// TIA Portal V20 export
// export: Created 2026-10-12T05:42:35.0167656Z, ExportSetting WithDefaults, DisplayName Totally Integrated Automation Portal, DisplayVersion V20, DisplayName TIA Portal Openness, DisplayVersion V20, DisplayName TIA Portal Teamcenter Gateway, DisplayVersion V20, DisplayName TIA Portal Version Control Interface, DisplayVersion V20, DisplayName SINAMICS Startdrive Advanced, DisplayVersion V20 SP1 Update 2, DisplayName SINAMICS Startdrive G110M, G120, G120C, G120D, G120P, G115D, DisplayVersion V20 SP1 Update 2, DisplayName SINAMICS Startdrive G130, G150, S120, S150, SINAMICS MV, G220, S200, S210, DisplayVersion V20 SP1 Update 2, DisplayName STEP 7 Professional, DisplayVersion V20, DisplayName STEP 7 Safety, DisplayVersion V20, DisplayName WinCC Basic/Comfort/Advanced, DisplayVersion V20, DisplayName WinCC Professional, DisplayVersion V20, DisplayName WinCC Unified, DisplayVersion V20
FUNCTION_BLOCK "FB_LD_PressDemoHome"   // FB7, LAD
{ S7_Optimized_Access := 'TRUE' }
VERSION : 0.1
// stored: AutoNumber true, IsIECCheckEnabled false, IsRetainMemResEnabled false, MemoryReserve 100, SetENOAutomatically false, UDAEnableTagReadback false
   VAR_INPUT
      Run { ExternalWritable := 'False'} : Bool;
      Reset { ExternalWritable := 'False'} : Bool;
      OwnerIndex { ExternalWritable := 'False'} : DInt;
      Delta { ExternalWritable := 'False'} : Time;
   END_VAR
   VAR_IN_OUT
      PressRam : "FB_CylinderCM";
      Door : "FB_CylinderCM";
      PartSlide : "FB_CylinderCM";
   END_VAR
   VAR
      Seq { ExternalWritable := 'False'} : "FRK_SequenceCtx";
      Row1 { ExternalWritable := 'False'} : "FRK_SequenceRow";
      Row2 { ExternalWritable := 'False'} : "FRK_SequenceRow";
      Row3 { ExternalWritable := 'False'} : "FRK_SequenceRow";
      Row4 { ExternalWritable := 'False'} : "FRK_SequenceRow";
      At0 { ExternalAccessible := 'False'; ExternalVisible := 'False'; ExternalWritable := 'False'} : Bool;
      At900 { ExternalAccessible := 'False'; ExternalVisible := 'False'; ExternalWritable := 'False'} : Bool;
      At910 { ExternalAccessible := 'False'; ExternalVisible := 'False'; ExternalWritable := 'False'} : Bool;
      At999 { ExternalAccessible := 'False'; ExternalVisible := 'False'; ExternalWritable := 'False'} : Bool;
      Ready1 { ExternalAccessible := 'False'; ExternalVisible := 'False'; ExternalWritable := 'False'} : Bool;
      Ready2 { ExternalAccessible := 'False'; ExternalVisible := 'False'; ExternalWritable := 'False'} : Bool;
      Ready3 { ExternalAccessible := 'False'; ExternalVisible := 'False'; ExternalWritable := 'False'} : Bool;
      Ready4 { ExternalAccessible := 'False'; ExternalVisible := 'False'; ExternalWritable := 'False'} : Bool;
      Ready5 { ExternalAccessible := 'False'; ExternalVisible := 'False'; ExternalWritable := 'False'} : Bool;
      Advance { ExternalAccessible := 'False'; ExternalVisible := 'False'; ExternalWritable := 'False'} : Bool;
   END_VAR
BEGIN

REGION Network 1
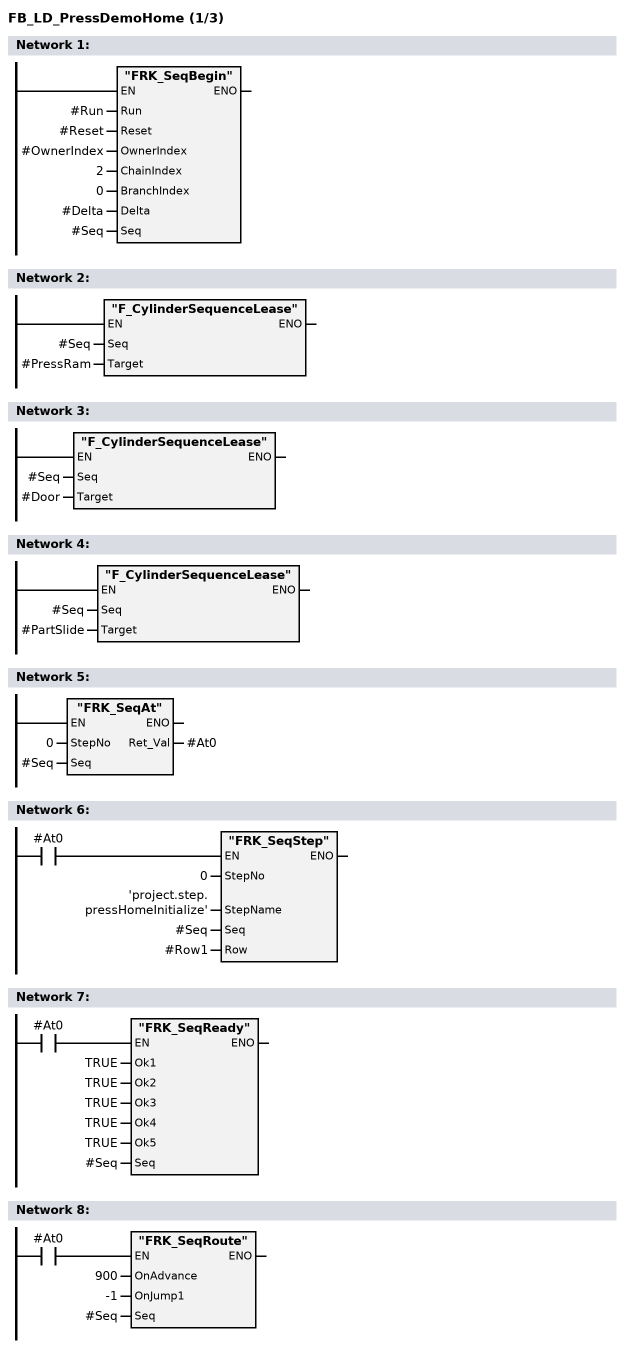
   RUNG wire#powerrail
      "FRK_SeqBegin"(Run := #Run, Reset := #Reset, OwnerIndex := #OwnerIndex, ChainIndex := 2, BranchIndex := 0, Delta := #Delta, Seq := #Seq)
   END_RUNG
   // the same network as SCL:
   "FRK_SeqBegin"(Run := #Run,
                  Reset := #Reset,
                  OwnerIndex := #OwnerIndex,
                  ChainIndex := 2,
                  BranchIndex := 0,
                  Delta := #Delta,
                  Seq := #Seq);
END_REGION

REGION Network 2
   RUNG wire#powerrail
      "F_CylinderSequenceLease"(Seq := #Seq, Target := #PressRam)
   END_RUNG
   // the same network as SCL:
   "F_CylinderSequenceLease"(Seq := #Seq, Target := #PressRam);
END_REGION

REGION Network 3
   RUNG wire#powerrail
      "F_CylinderSequenceLease"(Seq := #Seq, Target := #Door)
   END_RUNG
   // the same network as SCL:
   "F_CylinderSequenceLease"(Seq := #Seq, Target := #Door);
END_REGION

REGION Network 4
   RUNG wire#powerrail
      "F_CylinderSequenceLease"(Seq := #Seq, Target := #PartSlide)
   END_RUNG
   // the same network as SCL:
   "F_CylinderSequenceLease"(Seq := #Seq, Target := #PartSlide);
END_REGION

REGION Network 5
   RUNG wire#powerrail
      "FRK_SeqAt"(StepNo := 0, Seq := #Seq, Ret_Val => #At0)
   END_RUNG
   // the same network as SCL:
   #At0 := "FRK_SeqAt"(StepNo := 0, Seq := #Seq);
END_REGION

REGION Network 6
   RUNG wire#powerrail
      Contact( #At0 )
      "FRK_SeqStep"(StepNo := 0, StepName := 'project.step.pressHomeInitialize', Seq := #Seq, Row := #Row1)
   END_RUNG
   // the same network as SCL:
   IF #At0 THEN
       "FRK_SeqStep"(StepNo := 0, StepName := 'project.step.pressHomeInitialize', Seq := #Seq, Row := #Row1);
   END_IF;
END_REGION

REGION Network 7
   RUNG wire#powerrail
      Contact( #At0 )
      "FRK_SeqReady"(Ok1 := TRUE, Ok2 := TRUE, Ok3 := TRUE, Ok4 := TRUE, Ok5 := TRUE, Seq := #Seq)
   END_RUNG
   // the same network as SCL:
   IF #At0 THEN
       "FRK_SeqReady"(Ok1 := TRUE, Ok2 := TRUE, Ok3 := TRUE, Ok4 := TRUE, Ok5 := TRUE, Seq := #Seq);
   END_IF;
END_REGION

REGION Network 8
   RUNG wire#powerrail
      Contact( #At0 )
      "FRK_SeqRoute"(OnAdvance := 900, OnJump1 := -1, Seq := #Seq)
   END_RUNG
   // the same network as SCL:
   IF #At0 THEN "FRK_SeqRoute"(OnAdvance := 900, OnJump1 := -1, Seq := #Seq); END_IF;
END_REGION

REGION Network 9
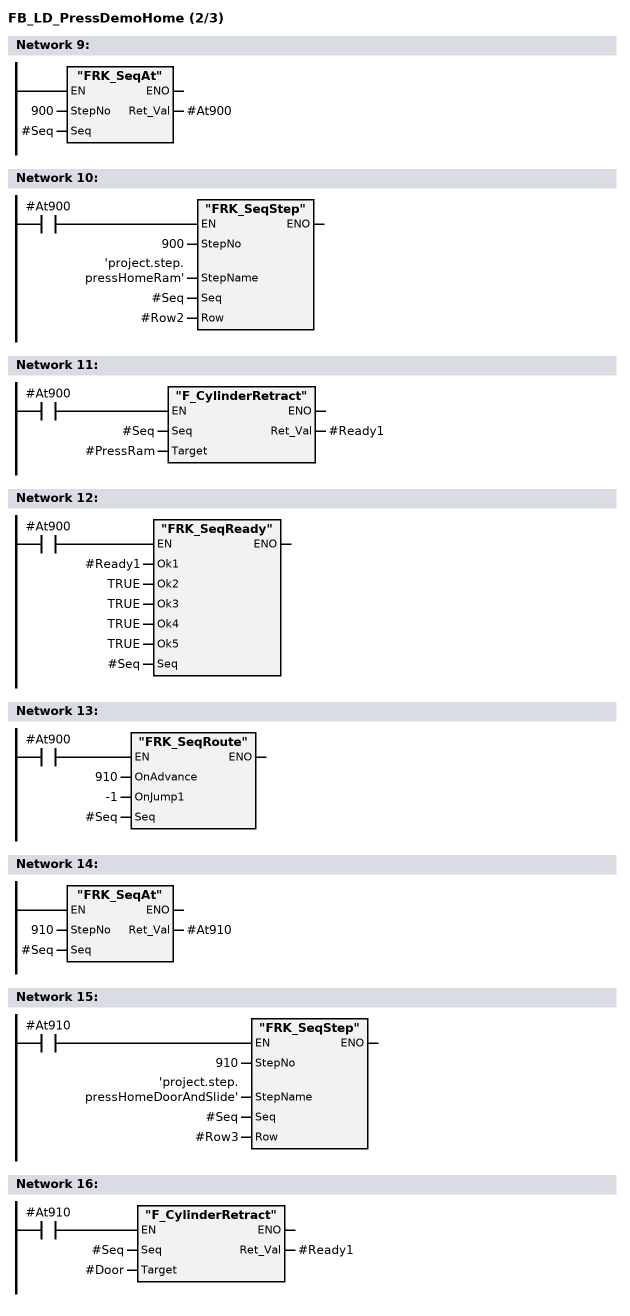
   RUNG wire#powerrail
      "FRK_SeqAt"(StepNo := 900, Seq := #Seq, Ret_Val => #At900)
   END_RUNG
   // the same network as SCL:
   #At900 := "FRK_SeqAt"(StepNo := 900, Seq := #Seq);
END_REGION

REGION Network 10
   RUNG wire#powerrail
      Contact( #At900 )
      "FRK_SeqStep"(StepNo := 900, StepName := 'project.step.pressHomeRam', Seq := #Seq, Row := #Row2)
   END_RUNG
   // the same network as SCL:
   IF #At900 THEN
       "FRK_SeqStep"(StepNo := 900, StepName := 'project.step.pressHomeRam', Seq := #Seq, Row := #Row2);
   END_IF;
END_REGION

REGION Network 11
   RUNG wire#powerrail
      Contact( #At900 )
      "F_CylinderRetract"(Seq := #Seq, Target := #PressRam, Ret_Val => #Ready1)
   END_RUNG
   // the same network as SCL:
   IF #At900 THEN #Ready1 := "F_CylinderRetract"(Seq := #Seq, Target := #PressRam); END_IF;
END_REGION

REGION Network 12
   RUNG wire#powerrail
      Contact( #At900 )
      "FRK_SeqReady"(Ok1 := #Ready1, Ok2 := TRUE, Ok3 := TRUE, Ok4 := TRUE, Ok5 := TRUE, Seq := #Seq)
   END_RUNG
   // the same network as SCL:
   IF #At900 THEN
       "FRK_SeqReady"(Ok1 := #Ready1, Ok2 := TRUE, Ok3 := TRUE, Ok4 := TRUE, Ok5 := TRUE, Seq := #Seq);
   END_IF;
END_REGION

REGION Network 13
   RUNG wire#powerrail
      Contact( #At900 )
      "FRK_SeqRoute"(OnAdvance := 910, OnJump1 := -1, Seq := #Seq)
   END_RUNG
   // the same network as SCL:
   IF #At900 THEN "FRK_SeqRoute"(OnAdvance := 910, OnJump1 := -1, Seq := #Seq); END_IF;
END_REGION

REGION Network 14
   RUNG wire#powerrail
      "FRK_SeqAt"(StepNo := 910, Seq := #Seq, Ret_Val => #At910)
   END_RUNG
   // the same network as SCL:
   #At910 := "FRK_SeqAt"(StepNo := 910, Seq := #Seq);
END_REGION

REGION Network 15
   RUNG wire#powerrail
      Contact( #At910 )
      "FRK_SeqStep"(StepNo := 910, StepName := 'project.step.pressHomeDoorAndSlide', Seq := #Seq, Row := #Row3)
   END_RUNG
   // the same network as SCL:
   IF #At910 THEN
       "FRK_SeqStep"(StepNo := 910, StepName := 'project.step.pressHomeDoorAndSlide', Seq := #Seq, Row := #Row3);
   END_IF;
END_REGION

REGION Network 16
   RUNG wire#powerrail
      Contact( #At910 )
      "F_CylinderRetract"(Seq := #Seq, Target := #Door, Ret_Val => #Ready1)
   END_RUNG
   // the same network as SCL:
   IF #At910 THEN #Ready1 := "F_CylinderRetract"(Seq := #Seq, Target := #Door); END_IF;
END_REGION

REGION Network 17
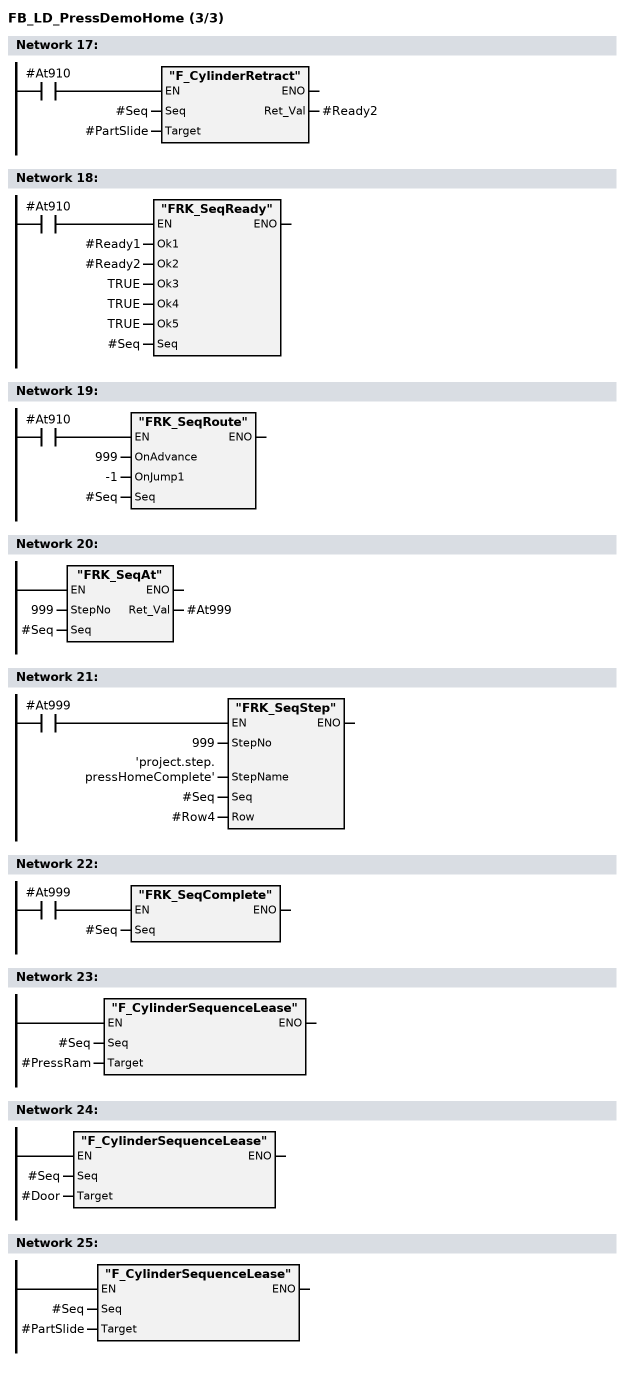
   RUNG wire#powerrail
      Contact( #At910 )
      "F_CylinderRetract"(Seq := #Seq, Target := #PartSlide, Ret_Val => #Ready2)
   END_RUNG
   // the same network as SCL:
   IF #At910 THEN #Ready2 := "F_CylinderRetract"(Seq := #Seq, Target := #PartSlide); END_IF;
END_REGION

REGION Network 18
   RUNG wire#powerrail
      Contact( #At910 )
      "FRK_SeqReady"(Ok1 := #Ready1, Ok2 := #Ready2, Ok3 := TRUE, Ok4 := TRUE, Ok5 := TRUE, Seq := #Seq)
   END_RUNG
   // the same network as SCL:
   IF #At910 THEN
       "FRK_SeqReady"(Ok1 := #Ready1, Ok2 := #Ready2, Ok3 := TRUE, Ok4 := TRUE, Ok5 := TRUE, Seq := #Seq);
   END_IF;
END_REGION

REGION Network 19
   RUNG wire#powerrail
      Contact( #At910 )
      "FRK_SeqRoute"(OnAdvance := 999, OnJump1 := -1, Seq := #Seq)
   END_RUNG
   // the same network as SCL:
   IF #At910 THEN "FRK_SeqRoute"(OnAdvance := 999, OnJump1 := -1, Seq := #Seq); END_IF;
END_REGION

REGION Network 20
   RUNG wire#powerrail
      "FRK_SeqAt"(StepNo := 999, Seq := #Seq, Ret_Val => #At999)
   END_RUNG
   // the same network as SCL:
   #At999 := "FRK_SeqAt"(StepNo := 999, Seq := #Seq);
END_REGION

REGION Network 21
   RUNG wire#powerrail
      Contact( #At999 )
      "FRK_SeqStep"(StepNo := 999, StepName := 'project.step.pressHomeComplete', Seq := #Seq, Row := #Row4)
   END_RUNG
   // the same network as SCL:
   IF #At999 THEN
       "FRK_SeqStep"(StepNo := 999, StepName := 'project.step.pressHomeComplete', Seq := #Seq, Row := #Row4);
   END_IF;
END_REGION

REGION Network 22
   RUNG wire#powerrail
      Contact( #At999 )
      "FRK_SeqComplete"(Seq := #Seq)
   END_RUNG
   // the same network as SCL:
   IF #At999 THEN "FRK_SeqComplete"(Seq := #Seq); END_IF;
END_REGION

REGION Network 23
   RUNG wire#powerrail
      "F_CylinderSequenceLease"(Seq := #Seq, Target := #PressRam)
   END_RUNG
   // the same network as SCL:
   "F_CylinderSequenceLease"(Seq := #Seq, Target := #PressRam);
END_REGION

REGION Network 24
   RUNG wire#powerrail
      "F_CylinderSequenceLease"(Seq := #Seq, Target := #Door)
   END_RUNG
   // the same network as SCL:
   "F_CylinderSequenceLease"(Seq := #Seq, Target := #Door);
END_REGION

REGION Network 25
   RUNG wire#powerrail
      "F_CylinderSequenceLease"(Seq := #Seq, Target := #PartSlide)
   END_RUNG
   // the same network as SCL:
   "F_CylinderSequenceLease"(Seq := #Seq, Target := #PartSlide);
END_REGION
END_FUNCTION_BLOCK
